Yaskawa INFORM job: TGTPROG.JBI

/JOB
//NAME TGTPROG
//POS
///NPOS 3,0,3,0,0,0
///TOOL 9
///POSTYPE PULSE
///PULSE
C00000=10000,-40000,-160000
C00001=500,-500,6000
C00002=-400,1200,10000
EC00000=9015
EC00001=3756
EC00002=-45150
//INST
<volatile>
///COMM Generated using RoboDK
///ATTR SC,RW
///GROUP1 RB1
NOP
'Program generated by RoboDK v
'6.0.7 for Yaskawa Motoman SCA
'RA on XX/XX/XXXX 18:00:00
'Using nominal kinematics.
MOVJ C00000 VJ=50.00  +MOVJ EC00000 VJ=100.00
MOVL C00001 V=100.0  +MOVJ EC00001 VJ=100.00
MOVJ C00002 VJ=50.00  +MOVJ EC00002 VJ=100.00
END
